Staubli VAL3: SpeedProg.pjx

--- SpeedProg.pjx ---
Parameters version=s7.5.3 stackSize=5000 millimeterUnit=true
Program file=MoveJoint.pgx
Program file=MoveLine.pgx
Program file=start.pgx
Program file=stop.pgx
Program file=main.pgx
Data file=SpeedProg.dtx

--- SpeedProg.dtx ---
mdesc mNomSpeed
frame fFrame1 = {x=1234.570, y=-98.765, z=50.500, rx=-0.000, ry=0.000, rz=30.000, fatherId=world[0]}
dio Input[16]
  [0] = {link=BasicIO-1\%I0}
  [1] = {link=BasicIO-1\%I1}
  [2] = {link=BasicIO-1\%I2}
  [3] = {link=BasicIO-1\%I3}
  [4] = {link=BasicIO-1\%I4}
  [5] = {link=BasicIO-1\%I5}
  [6] = {link=BasicIO-1\%I6}
  [7] = {link=BasicIO-1\%I7}
  [8] = {link=BasicIO-1\%I8}
  [9] = {link=BasicIO-1\%I9}
  [10] = {link=BasicIO-1\%I10}
  [11] = {link=BasicIO-1\%I11}
  [12] = {link=BasicIO-1\%I12}
  [13] = {link=BasicIO-1\%I13}
  [14] = {link=BasicIO-1\%I14}
  [15] = {link=BasicIO-1\%I15}
dio Output[16]
  [0] = {link=BasicIO-1\%Q0}
  [1] = {link=BasicIO-1\%Q1}
  [2] = {link=BasicIO-1\%Q2}
  [3] = {link=BasicIO-1\%Q3}
  [4] = {link=BasicIO-1\%Q4}
  [5] = {link=BasicIO-1\%Q5}
  [6] = {link=BasicIO-1\%Q6}
  [7] = {link=BasicIO-1\%Q7}
  [8] = {link=BasicIO-1\%Q8}
  [9] = {link=BasicIO-1\%Q9}
  [10] = {link=BasicIO-1\%Q10}
  [11] = {link=BasicIO-1\%Q11}
  [12] = {link=BasicIO-1\%Q12}
  [13] = {link=BasicIO-1\%Q13}
  [14] = {link=BasicIO-1\%Q14}
  [15] = {link=BasicIO-1\%Q15}
tool tCurrentTool = {x=10.000, y=20.000, z=150.000, rx=-0.000, ry=0.000, rz=-0.000, fatherId=flange[0], ioLink=ValveIO/valve1}
mdesc mCurrentSpeed
pointRs pPointRs = {fatherId=fFrame1[0]}
pointRs pPointRs2 = {fatherId=fFrame1[0]}

--- main.pgx ---
program main()
begin
  close(tCurrentTool)
  pPointRs.config.shoulder = lefty
  pPointRs2.config.shoulder = lefty
  mCurrentSpeed.tvel = 100.00
  mCurrentSpeed.blend = joint
  mCurrentSpeed.reach = 0.010
  mCurrentSpeed.leave = 0.010
  // Program SpeedProg start
  // Program generated by RoboDK v6.0.7 for Staubli TS20 FL 100 TC on XX/XX/XXXX 18:00:00
  // Using nominal kinematics.
  mCurrentSpeed.reach = 0.300
  mCurrentSpeed.leave = 0.300
  mCurrentSpeed.tvel = 1.000
  call MoveLine(-607.850,543.849,363.215,136.262,30.757,-130.375)
  call MoveJoint(10.00000,-20.00000,50.00000,30.00000)
  mCurrentSpeed.reach = 1.000
  mCurrentSpeed.leave = 1.000
  mCurrentSpeed.tvel = 12.300
  call MoveLine(-640.584,506.980,371.534,136.262,30.757,-130.375)
  call MoveJoint(30.00000,25.00000,80.00000,-45.00000)
  mCurrentSpeed.reach = 2.500
  mCurrentSpeed.leave = 2.500
  mCurrentSpeed.tvel = 99.900
  call MoveLine(-607.850,543.849,363.215,136.262,30.757,-130.375)
  call MoveJoint(10.00000,-20.00000,50.00000,30.00000)
  mCurrentSpeed.reach = 3.700
  mCurrentSpeed.leave = 3.700
  mCurrentSpeed.tvel = 333.333
  call MoveLine(-640.584,506.980,371.534,136.262,30.757,-130.375)
  call MoveJoint(30.00000,25.00000,80.00000,-45.00000)
  mCurrentSpeed.reach = 6.000
  mCurrentSpeed.leave = 6.000
  mCurrentSpeed.tvel = 1000.000
  call MoveLine(-607.850,543.849,363.215,136.262,30.757,-130.375)
  call MoveJoint(10.00000,-20.00000,50.00000,30.00000)
  mCurrentSpeed.reach = 9.000
  mCurrentSpeed.leave = 9.000
  mCurrentSpeed.tvel = 2500.000
  call MoveLine(-640.584,506.980,371.534,136.262,30.757,-130.375)
  call MoveJoint(30.00000,25.00000,80.00000,-45.00000)
  mCurrentSpeed.reach = 15.000
  mCurrentSpeed.leave = 15.000
  mCurrentSpeed.tvel = 5000.000
  call MoveLine(-607.850,543.849,363.215,136.262,30.757,-130.375)
  call MoveJoint(10.00000,-20.00000,50.00000,30.00000)
  mCurrentSpeed.reach = 30.000
  mCurrentSpeed.leave = 30.000
  mCurrentSpeed.tvel = 12000.000
  call MoveLine(-640.584,506.980,371.534,136.262,30.757,-130.375)
  call MoveJoint(30.00000,25.00000,80.00000,-45.00000)
  mCurrentSpeed.reach = 75.000
  mCurrentSpeed.leave = 75.000
  mCurrentSpeed.tvel = 0.500
  call MoveLine(-607.850,543.849,363.215,136.262,30.757,-130.375)
  call MoveJoint(10.00000,-20.00000,50.00000,30.00000)
  mCurrentSpeed.reach = 150.000
  mCurrentSpeed.leave = 150.000
  mCurrentSpeed.tvel = 750.000
  call MoveLine(-640.584,506.980,371.534,136.262,30.757,-130.375)
  call MoveJoint(30.00000,25.00000,80.00000,-45.00000)
  call MoveLine(-640.584,506.980,371.534,136.262,30.757,-130.375)

  waitEndMove()
  // Program SpeedProg end

end

--- start.pgx ---
program start()
begin
  call main()
end

--- MoveJoint.pgx ---
program MoveJoint(num x_nJ1, num x_nJ2, num x_nJ3, num x_nJ4)
  local joint l_jJoint
begin
  l_jJoint.j1 = x_nJ1
  l_jJoint.j2 = x_nJ2
  l_jJoint.j3 = x_nJ3
  l_jJoint.j4 = x_nJ4
  movej(l_jJoint,tCurrentTool ,mCurrentSpeed)
end

--- MoveLine.pgx ---
program MoveLine(num x_nX, num x_nY, num x_nZ, num x_nRx, num x_nRy, num x_nRz)
begin
  pPointRs.trsf.x = x_nX
  pPointRs.trsf.y = x_nY
  pPointRs.trsf.z = x_nZ
  pPointRs.trsf.rx = x_nRx
  pPointRs.trsf.ry = x_nRy
  pPointRs.trsf.rz = x_nRz
  movel(pPointRs,tCurrentTool,mCurrentSpeed)
end

--- stop.pgx ---
program stop()
begin
end
